Fanuc KAREL source: KA00046.KL

PROGRAM KA00046
%NOLOCKGROUP
VAR
  SRC: STRING[80]
  DST: CONFIG
BEGIN
  SRC = 'A'
  DST = SRC
END KA00046
